// TIA Portal V20 export
// export: Created 2026-10-12T16:46:21.5161049Z, ExportSetting WithDefaults, DisplayName Totally Integrated Automation Portal, DisplayVersion V20 Update 6, DisplayName TIA Portal Openness, DisplayVersion V20 Update 6, DisplayName TIA Portal Version Control Interface, DisplayVersion V20 Update 6, DisplayName SINAMICS Startdrive Advanced, DisplayVersion V20 SP1 Update 2, DisplayName SINAMICS Startdrive G110M, G120, G120C, G120D, G120P, G115D, DisplayVersion V20 SP1 Update 2, DisplayName SINAMICS Startdrive G130, G150, S120, S150, SINAMICS MV, G220, S200, S210, DisplayVersion V20 SP1 Update 2, DisplayName STEP 7 Professional, DisplayVersion V20 Update 6, DisplayName STEP 7 Safety, DisplayVersion V20 Update 2, DisplayName WinCC Basic/Comfort/Advanced, DisplayVersion V20 Update 6, DisplayName WinCC Professional, DisplayVersion V20 Update 6, DisplayName WinCC Unified, DisplayVersion V20 Update 6
DATA_BLOCK "FB_Anlagensteuerung_DB"   // DB1
VERSION : 0.9
// stored: AutoNumber true, DBAccessibleFromOPCUA true, DBAccessibleFromWebserver true, InstanceOfName FB_Anlagensteuerung, InstanceOfType FB
"FB_Anlagensteuerung"
   // VAR_INPUT
   //    Blink_Takt : Bool;
   //    Clock_10Hz : Bool;
   //    Not_Halt_Aktiv : Bool;
   // END_VAR
   // VAR
   //    Auftragsmanager { S7_SetPoint := 'True'} : "FB_Auftragsmanager";
   //    Bad { S7_SetPoint := 'True'} : Array[1.."c_Anzahl_Bad"] of "FB_Bad";
   //    Heizung { S7_SetPoint := 'True'} : "FB_Heizungssteuerung";
   //    Blink_Zaehler : Int;
   //    M_10Hz_Alt : Bool;
   // END_VAR
BEGIN
END_DATA_BLOCK
